(****************************************************************************************************<br>
© Syntegon Group.<br>
All rights reserved, also regarding any disposal, exploitation, reproduction, editing, distribution,<br>
as well as in the event of applications for industrial property rights.<br>
*****************************************************************************************************<br>
DESCRIPTION:<br>
DEMO ONLY: Cartesian application (Y = 6500..7300). A Cartesian robot picks products from the Cartesian infeed,<br>
turns them by C = -90 deg, tilts them by A while lowering and places them onto the Cartesian outfeed, every second<br>
one on top of the one it put down before (following it along the belt). Its gripper<br>
is a cup in the middle with two jaws beside it. Called by P_VisuDemo.<br>
****************************************************************************************************)
PROGRAM P_VisuDemoCartesian
VAR
	fb_CartInfeed						: _FB_VisuConveyor;
	fb_CartOutfeed						: _FB_VisuConveyor;
	fb_Cartesian						: _FB_VisuCartesian;

	(* Conveyors *)
	lr_Dt								: LREAL;	// [s] cycle time
	udn_Seed							: UDINT := 45678;	// [-] pseudo random generator state
	lr_InfeedPosition					: LREAL;	// [mm] belt position of the Cartesian infeed
	lr_OutfeedPosition					: LREAL;	// [mm] belt position of the Cartesian outfeed
	lr_SinceSpawn						: LREAL;	// [s] since the last product
	BeltPose							: ST_VisuPose;
	LatchPose							: ST_VisuPlanarPose;
	CartPose							: ST_VisuPose;

	(* Cartesian robot: axis actual values, start above the infeed *)
	n_CartPhase							: INT;
	lr_CartX							: LREAL := 900;	// [mm]
	lr_CartY							: LREAL := 200;	// [mm]
	lr_CartZ							: LREAL := -200;	// [mm]
	lr_CartC							: LREAL;	// [deg]
	lr_CartA							: LREAL;	// [deg]
	lr_CartPickC						: LREAL;	// [deg] C that turns the gripper onto the current product
	lr_CartJaw							: LREAL := 120;	// [mm] jaw distance from the cup along the gripper's X
	b_CartGrip							: BOOL;
	udn_CartProduct						: UDINT;	// [-] product id on the Cartesian infeed
	udn_CartStackBase					: UDINT;	// [-] product on the outfeed the next one is stacked on, 0 = the next one becomes it
	b_CartStacking						: BOOL;	// the product carried now goes onto udn_CartStackBase
END_VAR
VAR CONSTANT
	(* Robot turned by -90 deg: X axis across the belts towards MCS -Y (outfeed under X = 100, infeed under
	   X = 900), Y axis along MCS +X from X = 1000. *)
	lr_CART_INFEED_Y					: LREAL := 6500;	// [mm]
	lr_CART_OUTFEED_Y					: LREAL := 7300;	// [mm]
	lr_CART_BELT_LENGTH					: LREAL := 3000;	// [mm]
	lr_CART_BELT_SPEED					: LREAL := 150;	// [mm/s]
	lr_CART_SPAWN_INTERVAL				: LREAL := 2.5;	// [s]
	lr_CART_X							: LREAL := 1000;	// [mm]
	lr_CART_Y							: LREAL := 7400;	// [mm]
	lr_CART_Z							: LREAL := 1540;	// [mm] Z = -550 puts the cup's grip point (A = 0) on the product top
	lr_CART_TOOL_LENGTH					: LREAL := 150;	// [mm] flange to the cup's grip point
	lr_CART_CUP_HEIGHT					: LREAL := 40;	// [mm]
	lr_CART_JAW_DIAMETER				: LREAL := 20;	// [mm]
	lr_CART_JAW_HEIGHT					: LREAL := 120;	// [mm]
	lr_CART_JAW_TOP						: LREAL := 60;	// [mm] jaw tops below the flange
	lr_CART_JAW_OPEN					: LREAL := 120;	// [mm]
	lr_CART_JAW_CLOSED					: LREAL := 70;	// [mm] closed on a 120 mm product
	lr_CART_JAW_SPEED					: LREAL := 300;	// [mm/s]
	lr_CART_RAIL_HEIGHT					: LREAL := 1200;	// [mm]
	lr_CART_X_OUTFEED					: LREAL := 100;	// [mm]
	lr_CART_X_INFEED					: LREAL := 900;	// [mm]
	lr_CART_Y_HOME						: LREAL := 200;	// [mm]
	lr_CART_Y_STACK_BASE				: LREAL := 300;	// [mm] a product the next one is stacked on is put down here
	lr_CART_Y_STACK_MAX				: LREAL := 900;	// [mm] beyond this no stacking: the product below would leave the reach
	lr_CART_Z_PICK						: LREAL := -550;	// [mm]
	lr_CART_Z_TRAVEL					: LREAL := -200;	// [mm]
	lr_CART_TILT						: LREAL := 20;	// [deg] A while lowering
	lr_CART_TURN						: LREAL := -90;	// [deg] C between pick and place
	lr_CART_XY_SPEED					: LREAL := 1500;	// [mm/s]
	lr_CART_Z_SPEED						: LREAL := 800;	// [mm/s]
	lr_CART_C_SPEED						: LREAL := 180;	// [deg/s]
	lr_CART_A_SPEED						: LREAL := 60;	// [deg/s]
	n_CART_IDLE							: INT := 0;
	n_CART_DESCEND						: INT := 1;
	n_CART_LIFT							: INT := 2;
	n_CART_TRANSFER						: INT := 3;
	n_CART_LOWER						: INT := 4;
	n_CART_STRAIGHTEN					: INT := 5;
	n_CART_RELEASE						: INT := 6;
	n_CART_RISE							: INT := 7;
END_VAR

lr_Dt := DEMO_GlobalVar.DEMO_lr_Dt;


(****************************************************************************************************)
(* REGISTRATION (idempotent, every cycle)                                                           *)
(****************************************************************************************************)
fb_CartInfeed.m_Register(vio_Manifest := GVL_Visu.stManifest, vi_udn_Id := 8, vi_str_Name := 'Cartesian infeed');
fb_CartOutfeed.m_Register(vio_Manifest := GVL_Visu.stManifest, vi_udn_Id := 9, vi_str_Name := 'Cartesian outfeed');
fb_Cartesian.m_Register(vio_Manifest := GVL_Visu.stManifest, vi_udn_Id := 40, vi_str_Name := 'Cartesian');


(****************************************************************************************************)
(* CONVEYORS (configuration idempotent, every cycle)                                                *)
(****************************************************************************************************)
BeltPose.fX := 0;
BeltPose.fY := lr_CART_INFEED_Y;
BeltPose.fZ := DEMO_GlobalConst.DEMO_lr_BELT_Z;
fb_CartInfeed.m_SetPose(vi_Pose := BeltPose);
fb_CartInfeed.m_Configure(vi_lr_Length := lr_CART_BELT_LENGTH,
	vi_lr_Width := DEMO_GlobalConst.DEMO_lr_BELT_WIDTH);
BeltPose.fY := lr_CART_OUTFEED_Y;
fb_CartOutfeed.m_SetPose(vi_Pose := BeltPose);
fb_CartOutfeed.m_Configure(vi_lr_Length := lr_CART_BELT_LENGTH,
	vi_lr_Width := DEMO_GlobalConst.DEMO_lr_BELT_WIDTH);
(* The infeed's belt coordinates count from the robot's Y = 0, 1000 mm behind the belt start. *)
fb_CartInfeed.m_SetOriginShift(vi_lr_X := lr_CART_X, vi_lr_Y := 0, vi_lr_Z := 0);
fb_CartInfeed.m_SetProductType(vi_udn_Id := 1, vi_lr_Length := DEMO_GlobalConst.DEMO_lr_PRODUCT_LENGTH,
	vi_lr_Width := DEMO_GlobalConst.DEMO_lr_PRODUCT_WIDTH, vi_lr_Height := DEMO_GlobalConst.DEMO_lr_PRODUCT_HEIGHT,
	vi_e_Shape := E_VisuProductShape.BOX, vi_lr_CornerRadius := 0);
fb_CartOutfeed.m_SetProductType(vi_udn_Id := 1, vi_lr_Length := DEMO_GlobalConst.DEMO_lr_PRODUCT_LENGTH,
	vi_lr_Width := DEMO_GlobalConst.DEMO_lr_PRODUCT_WIDTH, vi_lr_Height := DEMO_GlobalConst.DEMO_lr_PRODUCT_HEIGHT,
	vi_e_Shape := E_VisuProductShape.BOX, vi_lr_CornerRadius := 0);

(* Belt travel *)
lr_InfeedPosition := lr_InfeedPosition + lr_CART_BELT_SPEED * lr_Dt;
lr_OutfeedPosition := lr_OutfeedPosition + lr_CART_BELT_SPEED * lr_Dt;
fb_CartInfeed.m_SetBeltPosition(lr_InfeedPosition);
fb_CartOutfeed.m_SetBeltPosition(lr_OutfeedPosition);


(****************************************************************************************************)
(* PRODUCT INFEED: regular gaps, products turned                                                    *)
(****************************************************************************************************)
lr_SinceSpawn := lr_SinceSpawn + lr_Dt;
IF lr_SinceSpawn >= lr_CART_SPAWN_INTERVAL THEN
	lr_SinceSpawn := 0;
	udn_Seed := udn_Seed * 1103515245 + 12345;
	LatchPose.fX := 100;
	LatchPose.fY := lr_CART_INFEED_Y;
	LatchPose.fZ := DEMO_GlobalConst.DEMO_lr_BELT_Z;
	LatchPose.fRz := (UDINT_TO_LREAL((udn_Seed / 1000) MOD 1000) / 1000.0 - 0.5) * 60.0;
	IF fb_CartInfeed.m_LatchProduct(vi_udn_Id := DEMO_GlobalVar.DEMO_udn_NextId,
		vi_LatchPose := fb_CartInfeed.m_McsToBelt(vi_Pose := LatchPose),
		vi_udn_ProductType := 1, vi_lr_LatchBeltPosition := 0, vi_b_UseLatchBeltPosition := FALSE,
		vi_e_State := E_VisuProductState.DETECTED, vi_udn_ClientId := 0)
	THEN
		DEMO_GlobalVar.DEMO_udn_NextId := DEMO_GlobalVar.DEMO_udn_NextId + 1;
	END_IF
END_IF


(****************************************************************************************************)
(* CARTESIAN ROBOT                                                                                  *)
(****************************************************************************************************)
CartPose.fX := lr_CART_X;
CartPose.fY := lr_CART_Y;
CartPose.fZ := lr_CART_Z;
CartPose.fRz := -90;
fb_Cartesian.m_SetPose(vi_Pose := CartPose);
fb_Cartesian.m_Configure(vi_lr_XMin := 0, vi_lr_XMax := 1200, vi_lr_YMin := 0, vi_lr_YMax := 1000,
	vi_lr_ZMin := -600, vi_lr_ZMax := 0, vi_lr_RailHeight := lr_CART_RAIL_HEIGHT);
(* Limit area in the robot frame (flange coordinates): X only up to the infeed, Z not into the top 100 mm. *)
fb_Cartesian.m_SetLimitArea(vi_lr_XMin := 0, vi_lr_XMax := 1000, vi_lr_YMin := 0, vi_lr_YMax := 1000,
	vi_lr_ZMin := -600, vi_lr_ZMax := -100);
(* Around the flange and the gripper below it. *)
fb_Cartesian.m_SetTcpLimitArea(vi_lr_XMin := -80, vi_lr_XMax := 80, vi_lr_YMin := -80, vi_lr_YMax := 80,
	vi_lr_ZMin := -50, vi_lr_ZMax := 20);
(* A cup in the middle carries the product, two jaws close beside it. *)
fb_Cartesian.m_SetFinger(vi_un_Finger := 1, vi_lr_Diameter := DEMO_GlobalConst.DEMO_lr_CUP_DIAMETER,
	vi_lr_Height := lr_CART_CUP_HEIGHT);
fb_Cartesian.m_SetFinger(vi_un_Finger := 2, vi_lr_Diameter := lr_CART_JAW_DIAMETER, vi_lr_Height := lr_CART_JAW_HEIGHT);
fb_Cartesian.m_SetFinger(vi_un_Finger := 3, vi_lr_Diameter := lr_CART_JAW_DIAMETER, vi_lr_Height := lr_CART_JAW_HEIGHT);
fb_Cartesian.m_SetZone(vi_un_Zone := 1, vi_udn_ConveyorId := fb_CartInfeed.m_Id(),
	vi_lr_Start := 0, vi_lr_End := 1000, vi_lr_AllocationOffset := 0, vi_lr_CcsOffset := 0,
	vi_lr_StartY := 0, vi_lr_EndY := 0);
fb_Cartesian.m_SetZone(vi_un_Zone := 2, vi_udn_ConveyorId := fb_CartOutfeed.m_Id(),
	vi_lr_Start := lr_CART_X + lr_CART_Y_STACK_BASE - 100, vi_lr_End := lr_CART_X + lr_CART_Y_STACK_MAX + 100,
	vi_lr_AllocationOffset := 0, vi_lr_CcsOffset := lr_CART_X + (lr_CART_Y_STACK_BASE + lr_CART_Y_STACK_MAX) / 2,
	vi_lr_StartY := 0, vi_lr_EndY := 0);
m_Step();
fb_Cartesian.m_SetAxes(vi_lr_X := lr_CartX, vi_lr_Y := lr_CartY, vi_lr_Z := lr_CartZ, vi_b_GripperActive := b_CartGrip);

(* C and A turn and tilt the gripper below the flange; they show only through the finger poses. *)
lr_CartJaw := _FC_DemoApproach(lr_CartJaw, SEL(b_CartGrip, lr_CART_JAW_OPEN, lr_CART_JAW_CLOSED), lr_CART_JAW_SPEED * lr_Dt);
fb_Cartesian.m_SetFingerState(vi_un_Finger := 1,
	vi_Pose := m_Finger(vi_lr_OffsetX := 0, vi_lr_OffsetZ := -(lr_CART_TOOL_LENGTH - lr_CART_CUP_HEIGHT)),
	vi_b_Active := b_CartGrip);
fb_Cartesian.m_SetFingerState(vi_un_Finger := 2,
	vi_Pose := m_Finger(vi_lr_OffsetX := lr_CartJaw, vi_lr_OffsetZ := -lr_CART_JAW_TOP),
	vi_b_Active := b_CartGrip);
fb_Cartesian.m_SetFingerState(vi_un_Finger := 3,
	vi_Pose := m_Finger(vi_lr_OffsetX := -lr_CartJaw, vi_lr_OffsetZ := -lr_CART_JAW_TOP),
	vi_b_Active := b_CartGrip);


(****************************************************************************************************)
(* HOUSEKEEPING                                                                                     *)
(****************************************************************************************************)
fb_CartInfeed.m_RemoveProductsBeyond(lr_CART_BELT_LENGTH + DEMO_GlobalConst.DEMO_lr_REMOVE_BEYOND_END);
fb_CartOutfeed.m_RemoveProductsBeyond(lr_CART_BELT_LENGTH + DEMO_GlobalConst.DEMO_lr_REMOVE_BEYOND_END);

(****************************************************************************************************<br>
© Syntegon Group.<br>
All rights reserved, also regarding any disposal, exploitation, reproduction, editing, distribution,<br>
as well as in the event of applications for industrial property rights.<br>
*****************************************************************************************************<br>
DESCRIPTION:<br>
Pose of a Cartesian gripper finger, absolute in the MCS: the finger sits at (vi_lr_OffsetX, 0, vi_lr_OffsetZ) in<br>
the gripper, which is turned by C about Z and tilted by A about its own X below the flange. The robot is<br>
turned by -90 deg: local (x, y, z) is MCS (lr_CART_X + y, lr_CART_Y - x, lr_CART_Z + z).<br>
****************************************************************************************************)
METHOD PRIVATE m_Finger : ST_VisuPose
VAR_INPUT
	vi_lr_OffsetX						: LREAL;	// [mm] along the gripper's X
	vi_lr_OffsetZ						: LREAL;	// [mm] below the flange: negative
END_VAR
VAR
	lr_TempA							: LREAL;	// [rad]
	lr_TempC							: LREAL;	// [rad]
	lr_TempVx							: LREAL;	// [mm] offset in the robot frame
	lr_TempVy							: LREAL;	// [mm]
	lr_TempVz							: LREAL;	// [mm]
END_VAR
lr_TempA := lr_CartA * VISU_GlobalConst.VISU_lr_DEG_TO_RAD;
lr_TempC := lr_CartC * VISU_GlobalConst.VISU_lr_DEG_TO_RAD;
(* Rz(C) * Rx(A) * (x, 0, z) *)
lr_TempVx := vi_lr_OffsetX * COS(lr_TempC) + vi_lr_OffsetZ * SIN(lr_TempA) * SIN(lr_TempC);
lr_TempVy := vi_lr_OffsetX * SIN(lr_TempC) - vi_lr_OffsetZ * SIN(lr_TempA) * COS(lr_TempC);
lr_TempVz := vi_lr_OffsetZ * COS(lr_TempA);
m_Finger.fX := lr_CART_X + (lr_CartY + lr_TempVy);
m_Finger.fY := lr_CART_Y - (lr_CartX + lr_TempVx);
m_Finger.fZ := lr_CART_Z + (lr_CartZ + lr_TempVz);
m_Finger.fRx := lr_CartA;
m_Finger.fRy := 0;
m_Finger.fRz := -90 + lr_CartC;
END_METHOD

(****************************************************************************************************<br>
© Syntegon Group.<br>
All rights reserved, also regarding any disposal, exploitation, reproduction, editing, distribution,<br>
as well as in the event of applications for industrial property rights.<br>
*****************************************************************************************************<br>
DESCRIPTION:<br>
Moves the Cartesian robot's axes one cycle towards the goal, each with its own speed. TRUE once all are there.<br>
****************************************************************************************************)
METHOD PRIVATE m_Move : BOOL
VAR_INPUT
	vi_lr_X								: LREAL;	// [mm]
	vi_lr_Y								: LREAL;	// [mm]
	vi_lr_Z								: LREAL;	// [mm]
	vi_lr_C								: LREAL;	// [deg]
	vi_lr_A								: LREAL;	// [deg]
END_VAR
lr_CartX := _FC_DemoApproach(lr_CartX, vi_lr_X, lr_CART_XY_SPEED * lr_Dt);
lr_CartY := _FC_DemoApproach(lr_CartY, vi_lr_Y, lr_CART_XY_SPEED * lr_Dt);
lr_CartZ := _FC_DemoApproach(lr_CartZ, vi_lr_Z, lr_CART_Z_SPEED * lr_Dt);
lr_CartC := _FC_DemoApproach(lr_CartC, vi_lr_C, lr_CART_C_SPEED * lr_Dt);
lr_CartA := _FC_DemoApproach(lr_CartA, vi_lr_A, lr_CART_A_SPEED * lr_Dt);
(* _FC_DemoApproach lands exactly on the goal, so equality is safe. *)
m_Move := lr_CartX = vi_lr_X AND lr_CartY = vi_lr_Y AND lr_CartZ = vi_lr_Z AND lr_CartC = vi_lr_C AND lr_CartA = vi_lr_A;
END_METHOD

(****************************************************************************************************<br>
© Syntegon Group.<br>
All rights reserved, also regarding any disposal, exploitation, reproduction, editing, distribution,<br>
as well as in the event of applications for industrial property rights.<br>
*****************************************************************************************************<br>
DESCRIPTION:<br>
Cartesian robot: follows a product on the Cartesian infeed in Y with the gripper turned onto it (C), picks<br>
it, carries it across to the outfeed while turning it by a further -90 deg, tilts it by A while lowering,<br>
straightens it and places it. Every second product goes on top of the one put down before, following it along<br>
the outfeed, as long as that one is in reach; otherwise it is put down at lr_CART_Y_STACK_BASE and the next one<br>
is stacked on it.<br>
****************************************************************************************************)
METHOD PRIVATE m_Step : BOOL
VAR
	n_TempFound							: INT;
	un_TempScan							: UINT;
	b_TempHave							: BOOL;
	lr_TempProductY						: LREAL;	// [mm] robot Y of the current product: its MCS x relative to the robot origin
	TempProduct							: ST_VisuProduct;
	TempProductPose						: ST_VisuPlanarPose;
	TempPlacePose						: ST_VisuPlanarPose;
	TempStackProduct					: ST_VisuProduct;
	TempStackPose						: ST_VisuPlanarPose;
	n_TempStackIdx						: INT;
	b_TempStackFound					: BOOL;
	lr_TempStackY						: LREAL;	// [mm] robot Y of the product to stack on
	lr_TempPlaceY						: LREAL;	// [mm] robot Y to put the product down at
	lr_TempPlaceZ						: LREAL;	// [mm] robot Z to put it down at: one product higher when stacking
	udn_TempPlacedId					: UDINT;
END_VAR
(* Current product *)
b_TempHave := FALSE;
IF udn_CartProduct <> 0 THEN
	n_TempFound := fb_CartInfeed.m_FindProduct(udn_CartProduct);
	IF n_TempFound >= 0 THEN
		b_TempHave := fb_CartInfeed.m_GetProduct(vi_un_Index := INT_TO_UINT(n_TempFound), vo_Product => TempProduct,
			vo_Pose => TempProductPose);
		TempProductPose := fb_CartInfeed.m_BeltToMcs(vi_Pose := TempProductPose);
		lr_TempProductY := TempProductPose.fX - lr_CART_X;
	END_IF
END_IF

(* Product to stack on, while it travels on the outfeed *)
b_TempStackFound := FALSE;
IF udn_CartStackBase <> 0 THEN
	n_TempStackIdx := fb_CartOutfeed.m_FindProduct(udn_CartStackBase);
	IF n_TempStackIdx >= 0 THEN
		fb_CartOutfeed.m_GetProduct(vi_un_Index := INT_TO_UINT(n_TempStackIdx), vo_Product => TempStackProduct,
			vo_Pose => TempStackPose);
		TempStackPose := fb_CartOutfeed.m_BeltToMcs(vi_Pose := TempStackPose);
		lr_TempStackY := TempStackPose.fX - lr_CART_X;
		b_TempStackFound := TRUE;
	END_IF
END_IF
IF NOT b_TempStackFound THEN
	b_CartStacking := FALSE;
END_IF
lr_TempPlaceY := SEL(b_CartStacking, lr_CART_Y_STACK_BASE, lr_TempStackY);
lr_TempPlaceZ := lr_CART_Z_PICK + SEL(b_CartStacking, 0, DEMO_GlobalConst.DEMO_lr_PRODUCT_HEIGHT);

(* Sequence *)
CASE n_CartPhase OF
	n_CART_IDLE:
		un_TempScan := 0;
		WHILE udn_CartProduct = 0 AND un_TempScan < fb_CartInfeed.m_ProductCount() DO
			fb_CartInfeed.m_GetProduct(vi_un_Index := un_TempScan, vo_Product => TempProduct, vo_Pose => TempProductPose);
			TempProductPose := fb_CartInfeed.m_BeltToMcs(vi_Pose := TempProductPose);
			IF TempProduct.eState = E_VisuProductState.DETECTED
			AND TempProductPose.fX - lr_CART_X >= 100
			AND TempProductPose.fX - lr_CART_X <= 600
			THEN
				fb_CartInfeed.m_SetProductState(vi_udn_Id := TempProduct.nId, vi_e_State := E_VisuProductState.ASSIGNED,
					vi_udn_ClientId := fb_Cartesian.m_Id(), vi_udn_MoverId := 0, vi_udn_FingerId := 0);
				udn_CartProduct := TempProduct.nId;
				(* The gripper's +X in the MCS is pose rz (-90 deg) + C. *)
				lr_CartPickC := TempProductPose.fRz + 90;
				n_CartPhase := n_CART_DESCEND;
			END_IF
			un_TempScan := un_TempScan + 1;
		END_WHILE
		IF udn_CartProduct = 0 THEN
			m_Move(vi_lr_X := lr_CART_X_INFEED, vi_lr_Y := lr_CART_Y_HOME, vi_lr_Z := lr_CART_Z_TRAVEL, vi_lr_C := 0,
				vi_lr_A := 0);
		END_IF

	n_CART_DESCEND:
		IF NOT b_TempHave THEN
			udn_CartProduct := 0;
			n_CartPhase := n_CART_RISE;
		ELSIF lr_TempProductY > 1000 THEN
			(* Out of reach: hand it back, it will be missed. *)
			fb_CartInfeed.m_SetProductState(vi_udn_Id := udn_CartProduct, vi_e_State := E_VisuProductState.DETECTED,
				vi_udn_ClientId := fb_Cartesian.m_Id(), vi_udn_MoverId := 0, vi_udn_FingerId := 0);
			udn_CartProduct := 0;
			n_CartPhase := n_CART_RISE;
		ELSIF m_Move(vi_lr_X := lr_CART_X_INFEED, vi_lr_Y := lr_TempProductY, vi_lr_Z := lr_CartZ,
			vi_lr_C := lr_CartPickC, vi_lr_A := 0)
		THEN
			(* Lowers only once above the product with the gripper turned onto it. *)
			IF m_Move(vi_lr_X := lr_CART_X_INFEED, vi_lr_Y := lr_TempProductY, vi_lr_Z := lr_CART_Z_PICK,
				vi_lr_C := lr_CartPickC, vi_lr_A := 0)
			THEN
				fb_CartInfeed.m_SetProductState(vi_udn_Id := udn_CartProduct, vi_e_State := E_VisuProductState.PICKED,
					vi_udn_ClientId := fb_Cartesian.m_Id(), vi_udn_MoverId := 0, vi_udn_FingerId := 1);
				b_CartGrip := TRUE;
				n_CartPhase := n_CART_LIFT;
			END_IF
		END_IF

	n_CART_LIFT:
		IF m_Move(vi_lr_X := lr_CartX, vi_lr_Y := lr_CartY, vi_lr_Z := lr_CART_Z_TRAVEL, vi_lr_C := lr_CartC,
			vi_lr_A := lr_CartA)
		THEN
			n_CartPhase := n_CART_TRANSFER;
		END_IF

	n_CART_TRANSFER:
		(* Every second product goes onto the one put down before, as long as that one is in reach. *)
		b_CartStacking := b_TempStackFound AND lr_TempStackY <= lr_CART_Y_STACK_MAX;
		IF NOT b_CartStacking THEN
			udn_CartStackBase := 0;
		END_IF
		lr_TempPlaceY := SEL(b_CartStacking, lr_CART_Y_STACK_BASE, lr_TempStackY);
		lr_TempPlaceZ := lr_CART_Z_PICK + SEL(b_CartStacking, 0, DEMO_GlobalConst.DEMO_lr_PRODUCT_HEIGHT);
		IF m_Move(vi_lr_X := lr_CART_X_OUTFEED, vi_lr_Y := lr_TempPlaceY, vi_lr_Z := lr_CART_Z_TRAVEL,
			vi_lr_C := lr_CartPickC + lr_CART_TURN, vi_lr_A := 0)
		THEN
			n_CartPhase := n_CART_LOWER;
		END_IF

	n_CART_LOWER:
		IF m_Move(vi_lr_X := lr_CartX, vi_lr_Y := lr_TempPlaceY, vi_lr_Z := lr_TempPlaceZ, vi_lr_C := lr_CartC,
			vi_lr_A := lr_CART_TILT)
		THEN
			n_CartPhase := n_CART_STRAIGHTEN;
		END_IF

	n_CART_STRAIGHTEN:
		IF m_Move(vi_lr_X := lr_CartX, vi_lr_Y := lr_TempPlaceY, vi_lr_Z := lr_CartZ, vi_lr_C := lr_CartC, vi_lr_A := 0) THEN
			n_CartPhase := n_CART_RELEASE;
		END_IF

	n_CART_RELEASE:
		(* Put down on the outfeed: it no longer lies on the infeed. *)
		fb_CartInfeed.m_RemoveProduct(udn_CartProduct);
		(* Turned by -90 deg: the cup (A = 0) is at MCS x = origin + Y, y = origin - X; the product keeps the turn. *)
		TempPlacePose.fX := lr_CART_X + lr_CartY;
		TempPlacePose.fY := lr_CART_Y - lr_CartX;
		(* A stacked product lies one product height above the belt. *)
		TempPlacePose.fZ := DEMO_GlobalConst.DEMO_lr_BELT_Z + SEL(b_CartStacking, 0, DEMO_GlobalConst.DEMO_lr_PRODUCT_HEIGHT);
		TempPlacePose.fRz := -90 + lr_CartC;
		udn_TempPlacedId := DEMO_GlobalVar.DEMO_udn_NextId;
		IF fb_CartOutfeed.m_LatchProduct(vi_udn_Id := DEMO_GlobalVar.DEMO_udn_NextId,
			vi_LatchPose := fb_CartOutfeed.m_McsToBelt(vi_Pose := TempPlacePose),
			vi_udn_ProductType := 1, vi_lr_LatchBeltPosition := 0, vi_b_UseLatchBeltPosition := FALSE,
			vi_e_State := E_VisuProductState.PLACED, vi_udn_ClientId := fb_Cartesian.m_Id())
		THEN
			DEMO_GlobalVar.DEMO_udn_NextId := DEMO_GlobalVar.DEMO_udn_NextId + 1;
		END_IF
		(* The next product goes onto this one, unless this one is already on top of another. *)
		IF b_CartStacking THEN
			udn_CartStackBase := 0;
		ELSE
			udn_CartStackBase := udn_TempPlacedId;
		END_IF
		b_CartStacking := FALSE;
		udn_CartProduct := 0;
		b_CartGrip := FALSE;
		n_CartPhase := n_CART_RISE;

	n_CART_RISE:
		IF m_Move(vi_lr_X := lr_CartX, vi_lr_Y := lr_CartY, vi_lr_Z := lr_CART_Z_TRAVEL, vi_lr_C := lr_CartC,
			vi_lr_A := lr_CartA)
		THEN
			n_CartPhase := n_CART_IDLE;
		END_IF
END_CASE
m_Step := TRUE;
END_METHOD

END_PROGRAM

(* stored: Version 1.1.0.1
   POU P_VisuDemoCartesian: Id {d5e22a24-ae42-4c62-9790-0f1f0f48b7a7}, SpecialFunc None
   Method m_Finger: Id {2e68f6f4-3124-4ca2-ba4d-f784a4bc7fa2}
   Method m_Move: Id {dce46312-c5f0-47a4-acbf-bc429aa07c03}
   Method m_Step: Id {05fd5b17-c85a-40bb-ba82-87c8709ed353} *)
